(* IEC 61131-3 sources: plc-process-lib/tests/POUs/Suites/FB_Runtime_Test, 14 files *)

(* ---- FB_Runtime_Test.decl.st ---- *)
// Назначение: набор зондов времени выполнения — вопросы раздела 24.2 контракта и ограничения
//             раздела 2.8, которые решает тест на CODESYS Control Win V3 (32 бит): монотонность и
//             разрешение LTIME() (по циклам задачи и внутри цикла), связывание вызова метода без
//             THIS^, частичный инициализатор массива структур, беззнаковая арифметика LTIME и
//             счётчиков, локальные экземпляры устройств в методе теста, цена копирования LKG.
//             Тест Runtime_LTime_MonotonicAcrossTaskCycles идёт 50 циклов задачи: его состояние —
//             в переменных набора (локальные переменные метода создаются заново каждый вызов).
// Автор:      kr0nsch
// Версия:     0.1.0
// Документ:   docs/TESTING.md, раздел «Зонды времени выполнения»
FUNCTION_BLOCK FB_Runtime_Test EXTENDS coUnit.FB_TestSuite
VAR CONSTANT
    RT_SAMPLES : UINT := 50;                       // циклов задачи в тесте по циклам
END_VAR
VAR
    fbRtSysTime : FB_SystemTime;                  // системное время для теста по циклам
    uiRtCount   : UINT;                           // записано отметок
    altRtStamp  : ARRAY[0..RT_SAMPLES - 1] OF LTIME;   // LTIME() в каждом цикле задачи
END_VAR

(* ---- CallDevice.method.decl.st ---- *)
// Помощник: вызов одного устройства массива со всеми VAR_IN_OUT (короче цикл теста)
METHOD PRIVATE CallDevice
VAR_IN_OUT
    fbDevice : FB_TestDeviceExt;    // устройство
    stCmdDev : ST_TestDeviceCmd;    // его команды
    stRetDev : ST_DeviceRetain;     // его retain
END_VAR
VAR_IN_OUT CONSTANT
    stCfgDev : ST_TestDeviceCfg;    // конфигурация
END_VAR
VAR_INPUT
    itfTimeSrc : I_TimeSource;      // источник времени
END_VAR

(* ---- LkgCopy300MotorCfgBelow1ms.method.decl.st ---- *)
// R13 контракта (данные для Control Win V3, не для ПЛК210): 300 копирований ST_MotorCfg (216 байт —
// копия LKG одного двигателя за цикл) занимают меньше 1 мс.
METHOD PRIVATE LkgCopy300MotorCfgBelow1ms
VAR
    fbSys   : FB_SystemTime;   // системное время
    stSrc   : ST_MotorCfg;     // источник копии
    stDst   : ST_MotorCfg;     // приёмник копии
    ltStart : LTIME;           // начало замера
    ltEnd   : LTIME;           // конец замера
    iStep   : INT;             // шаг цикла
END_VAR

(* ---- LkgCopy300MotorCfgBelow1ms.method.impl.st ---- *)
coUnit.TEST('Runtime_LkgCopy300MotorCfg_Below1ms');

ltStart := fbSys.Now();
FOR iStep := 1 TO 300 DO
    stSrc.tMinRun := INT_TO_TIME(iStep);
    stDst := stSrc;
END_FOR
ltEnd := fbSys.Now();
AssertEquals_TIME(Expected := T#300MS, Actual := stDst.tMinRun, Message := 'last copy done');
AssertTrue(Condition := ltEnd >= ltStart, Message := 'time does not decrease');
AssertTrue(Condition := ltEnd - ltStart < LTIME#1MS, Message := '300 copies of ST_MotorCfg below 1 ms');

coUnit.TEST_FINISHED();

(* ---- LocalDeviceInstancesRunInTestMethod.method.decl.st ---- *)
// R5 контракта: шесть экземпляров устройства (FB_TestDeviceExt: 8 слотов FB_Alarm, LKG) и их
// структуры — локальные переменные метода теста; стека задачи хватает, все работают.
METHOD PRIVATE LocalDeviceInstancesRunInTestMethod
VAR
    fbTime   : FB_FakeTime;                            // подменное время
    afbDev   : ARRAY[0..5] OF FB_TestDeviceExt;        // устройства в стеке метода
    astCmd   : ARRAY[0..5] OF ST_TestDeviceCmd;        // их команды
    astRet   : ARRAY[0..5] OF ST_DeviceRetain;         // их retain
    stCfg    : ST_TestDeviceCfg;                       // общая конфигурация
    itfDev   : I_Device;                               // устройство через интерфейс
    uiDev    : UINT;                                   // номер устройства
    xAllAuto : BOOL := TRUE;                           // все перешли в Auto
END_VAR

(* ---- LocalDeviceInstancesRunInTestMethod.method.impl.st ---- *)
coUnit.TEST('Runtime_LocalDeviceInstances_RunInTestMethod');

FOR uiDev := 0 TO 5 DO
    itfDev := afbDev[uiDev];
    itfDev.RequestMode(eNewMode := E_DeviceMode.Auto);
    CallDevice(fbDevice := afbDev[uiDev], stCmdDev := astCmd[uiDev], stRetDev := astRet[uiDev], stCfgDev := stCfg,
               itfTimeSrc := fbTime);
    xAllAuto := xAllAuto AND itfDev.Mode = E_DeviceMode.Auto;
END_FOR
AssertTrue(Condition := xAllAuto, Message := 'six local device instances run');

coUnit.TEST_FINISHED();

(* ---- LTimeMonotonicAcrossTaskCycles.method.decl.st ---- *)
// R1 контракта по циклам задачи: LTIME() (FB_SystemTime) в 50 циклах TestTask (10 мс) строго
// растёт от цикла к циклу, а промежуток 49 циклов — от 49·5 мс до 49·50 мс (время идёт с реальной
// скоростью). Единственный тест библиотеки на несколько циклов: реального ожидания в нём нет,
// цикл задачи — данность. Смену системного времени ОС тест не делает (нужны права администратора).
METHOD PRIVATE LTimeMonotonicAcrossTaskCycles
VAR
    uiIdx    : UINT;            // номер отметки
    xStrict  : BOOL := TRUE;    // каждая следующая отметка больше предыдущей
    ltSpan   : LTIME;           // от первой до последней отметки
END_VAR

(* ---- LTimeMonotonicAcrossTaskCycles.method.impl.st ---- *)
coUnit.TEST('Runtime_LTime_MonotonicAcrossTaskCycles');

IF uiRtCount < RT_SAMPLES THEN
    altRtStamp[uiRtCount] := fbRtSysTime.Now();
    uiRtCount := uiRtCount + 1;
ELSE
    FOR uiIdx := 1 TO RT_SAMPLES - 1 DO
        xStrict := xStrict AND (altRtStamp[uiIdx] > altRtStamp[uiIdx - 1]);
    END_FOR
    IF xStrict THEN
        ltSpan := altRtStamp[RT_SAMPLES - 1] - altRtStamp[0];
    ELSE
        ltSpan := LTIME#0S;
    END_IF
    AssertTrue(Condition := xStrict, Message := 'LTIME() strictly increases from task cycle to task cycle');
    AssertTrue(Condition := ltSpan >= LTIME#245MS, Message := '49 task cycles of 10 ms last at least 245 ms');
    AssertTrue(Condition := ltSpan <= LTIME#2S450MS, Message := '49 task cycles of 10 ms last at most 2.45 s');
    coUnit.TEST_FINISHED();
END_IF

(* ---- LTimeResolutionAtMost1us.method.decl.st ---- *)
// R1 контракта внутри цикла: 20 000 чтений LTIME() подряд — время не убывает, меняется хотя бы
// раз, наименьший ненулевой шаг (разрешение источника) не больше 1 мкс.
METHOD PRIVATE LTimeResolutionAtMost1us
VAR
    fbSys      : FB_SystemTime;     // источник под тестом
    itfTime    : I_TimeSource;      // через интерфейс, как в ФБ библиотеки
    ltPrev     : LTIME;             // предыдущее чтение
    ltNow      : LTIME;             // текущее чтение
    ltMinStep  : LTIME := LTIME#1S; // наименьший ненулевой шаг
    uiChanges  : UINT;              // сколько раз время изменилось
    xMonotonic : BOOL := TRUE;      // не убывало
    iStep      : INT;               // шаг цикла
END_VAR

(* ---- LTimeResolutionAtMost1us.method.impl.st ---- *)
coUnit.TEST('Runtime_LTime_ResolutionAtMost1us');

itfTime := fbSys;
ltPrev := itfTime.Now();
FOR iStep := 1 TO 20000 DO
    ltNow := itfTime.Now();
    xMonotonic := xMonotonic AND (ltNow >= ltPrev);
    IF ltNow > ltPrev THEN
        uiChanges := uiChanges + 1;
        IF ltNow - ltPrev < ltMinStep THEN
            ltMinStep := ltNow - ltPrev;
        END_IF
    END_IF
    ltPrev := ltNow;
END_FOR
AssertTrue(Condition := xMonotonic, Message := 'LTIME() does not decrease');
AssertTrue(Condition := uiChanges > 0, Message := 'LTIME() changes within 20000 reads');
AssertTrue(Condition := ltMinStep <= LTIME#1US, Message := 'smallest non-zero step at most 1 us');

coUnit.TEST_FINISHED();

(* ---- LTimeSubtractionWrapsWhenNegative.method.decl.st ---- *)
// L7 контракта: LTIME без знака — разность a - b при a < b не отрицательна, а переполняется по
// модулю 2^64 (огромное значение больше a), поэтому библиотека сравнивает отметки до вычитания.
METHOD PRIVATE LTimeSubtractionWrapsWhenNegative
VAR
    ltA : LTIME := LTIME#1S;   // меньшая отметка
    ltB : LTIME := LTIME#2S;   // большая отметка
    ltD : LTIME;               // a - b
END_VAR

(* ---- MethodCallWithoutThisDispatchesVirtually.method.decl.st ---- *)
// Связывание вызовов (L6 контракта): метод базы вызывает переопределённый метод через THIS^ и без
// него; у экземпляра наследника оба вызова выполняют реализацию наследника, у экземпляра базы —
// базы.
METHOD PRIVATE MethodCallWithoutThisDispatchesVirtually
VAR
    fbBase    : FB_ProbeHookBase;      // экземпляр базы
    fbDerived : FB_ProbeHookDerived;   // экземпляр наследника
END_VAR

(* ---- PartialArrayInitializerRestGetsElementDefaults.method.decl.st ---- *)
// R9 контракта: частичный инициализатор astAlarm в объявлении переменной Cfg (как в GVL_Persist)
// задаёт слот 0, остальные слоты получают умолчания ST_AlarmCfg (Medium), а не умолчания DUT
// устройства (у ST_AnalogInputCfg: слот 1 — Low, слот 3 — High); поля Cfg вне инициализатора
// сохраняют умолчания DUT.
METHOD PRIVATE PartialArrayInitializerRestGetsElementDefaults
VAR
    stPart : ST_AnalogInputCfg := (rRangeHi_eu := 5.0, astAlarm := [(ePriority := E_AlarmPriority.Low)]);   // зонд
    stFull : ST_AnalogInputCfg;   // умолчания DUT для сравнения
    stSlot : ST_AlarmCfg;         // копия слота
END_VAR

(* ---- UnsignedCountersWrapToZero.method.decl.st ---- *)
// Счётчики «по кругу» (uiCmdSeq, udiSeq): UINT 65535 + 1 и UDINT 4294967295 + 1 дают 0 без
// исключения на Control Win V3.
METHOD PRIVATE UnsignedCountersWrapToZero
VAR
    uiCnt  : UINT := 65535;         // счётчик UINT на пределе
    udiCnt : UDINT := 4294967295;   // счётчик UDINT на пределе
END_VAR
